(* IEC 61131-3 sources: RAG_PLC/data/result/test/009, 2 files *)

(* ---- wrapped.st ---- *)
(* =========================================================
   Generated by PLC-Eval Benchmark Wrapper
   ========================================================= *)

FUNCTION_BLOCK LLM_Wrapper_FB
VAR_INPUT
    SEP : BYTE;
END_VAR

VAR_IN_OUT
    LIST : oscat_STRING250;
END_VAR

VAR_OUTPUT
    LIST_CLEAN : BOOL;
END_VAR

VAR
    BUF_TO_STRING : BUF_TO_STRING;
    pt : oscat_bya_LIST_CLEAN;
    read : INT;
    write : INT := 1;
    last : BYTE;
    c : BYTE;
    cnt : INT;
    z : INT;
END_VAR

(*@KEY@: WORKSHEET
NAME: LIST_CLEAN
IEC_LANGUAGE: ST
*)
last := BYTE#0;
cnt := LEN(LIST);
write := 0;
FOR read := 1 TO cnt DO
    c := INT_TO_BYTE(GET_CHAR(LIST, read));
    IF c <> SEP OR last <> SEP THEN
        write := write + 1;
        pt[write] := c;
    END_IF;
    last := c;
END_FOR;
IF last = SEP THEN write := write - 1; END_IF;

FOR z := 0 TO 1 DO
    BUF_TO_STRING.REQ := z > 0;
    BUF_TO_STRING.BUF_FORMAT := TRUE;
    BUF_TO_STRING.BUF_OFFS := DINT#0;
    BUF_TO_STRING.BUF_CNT := INT_TO_DINT(write);
    BUF_TO_STRING.BUFFER := pt;
    BUF_TO_STRING.DST := LIST;
    BUF_TO_STRING();
    pt := BUF_TO_STRING.BUFFER;
    LIST := BUF_TO_STRING.DST;
END_FOR;

LIST_CLEAN := TRUE; (* 返回 TRUE *)
END_FUNCTION_BLOCK

PROGRAM Auto_Proxy_Prg
  VAR
    instance : LLM_Wrapper_FB;
  END_VAR

  instance();
END_PROGRAM

CONFIGURATION Config0
  RESOURCE Res0 ON PLC
    TASK TaskMain(INTERVAL := T#20ms, PRIORITY := 0);
    PROGRAM Inst0 WITH TaskMain : Auto_Proxy_Prg;
  END_RESOURCE
END_CONFIGURATION

(* ---- raw_code.st ---- *)
VAR_INPUT
    SEP : BYTE;
END_VAR

VAR_IN_OUT
    LIST : oscat_STRING250;
END_VAR

VAR_OUTPUT
    LIST_CLEAN : BOOL;
END_VAR

VAR
    BUF_TO_STRING : BUF_TO_STRING;
    pt : oscat_bya_LIST_CLEAN;
    read : INT;
    write : INT := 1;
    last : BYTE;
    c : BYTE;
    cnt : INT;
    z : INT;
END_VAR

(*@KEY@: WORKSHEET
NAME: LIST_CLEAN
IEC_LANGUAGE: ST
*)
last := BYTE#0;
cnt := LEN(LIST);
write := 0;
FOR read := 1 TO cnt DO
    c := INT_TO_BYTE(GET_CHAR(LIST, read));
    IF c <> SEP OR last <> SEP THEN
        write := write + 1;
        pt[write] := c;
    END_IF;
    last := c;
END_FOR;
IF last = SEP THEN write := write - 1; END_IF;

FOR z := 0 TO 1 DO
    BUF_TO_STRING.REQ := z > 0;
    BUF_TO_STRING.BUF_FORMAT := TRUE;
    BUF_TO_STRING.BUF_OFFS := DINT#0;
    BUF_TO_STRING.BUF_CNT := INT_TO_DINT(write);
    BUF_TO_STRING.BUFFER := pt;
    BUF_TO_STRING.DST := LIST;
    BUF_TO_STRING();
    pt := BUF_TO_STRING.BUFFER;
    LIST := BUF_TO_STRING.DST;
END_FOR;

LIST_CLEAN := TRUE; (* 返回 TRUE *)
